TYPE ST_ES_PB :
STRUCT
	in: BOOL;
	State: BOOL;
	Memo: BOOL;
	ByPass: BOOL;
	stBitMap                : STRING:= 'ImagePool.EStop_OK2'; //'ImagePool.EStop_ACT2'
END_STRUCT
END_TYPE

(* stored: Version 1.1.0.1, ProductVersion 3.1.4024.13
   DUT ST_ES_PB: Id {a16fcc2f-482c-4ee9-9b54-bbe315c0d3ca} *)
